(* IEC 61131-3 sources: SRCI_CLIENT_PLC/RobotLibrary/Library/POUs/Read/MC_ReadActualTCPVelocity/Structures, 4 files *)

(* ---- ReadActualTCPVelocityOutCmd.st ---- *)
{attribute 'pack_mode' := '1'}
// -------------------------------------------------------------------------
//  SRCI Robot Library
// -------------------------------------------------------------------------
//
//  Object:      ReadActualTCPVelocityOutCmd
//  Author:      Thorsten Brach
//  Date:        2024-08-09
//
//  Description:
//
//
//  Copyright:
//    (C) 2024 Thorsten Brach. All rights reserved
//             Licensed under the MIT License.
//
//  Disclaimer:
//    This project is provided without any guarantee and can be used for
//    private and commercial purposes. Any use is at the user’s
//    own risk and responsibility.
//
// -------------------------------------------------------------------------
TYPE ReadActualTCPVelocityOutCmd :
STRUCT
  /// Absolute actual velocity of the robot’s TCP. [mm/s]
  ActualTCPVelocity  : REAL;
  /// Index of tool of returned velocity
  /// •      0: Flange
  /// • 1..254: Tool frames
  ToolNoReturn       : USINT;
  /// Index of frame of returned position
  /// •      0: WCS
  /// • 1..254: User frames
  FrameNoReturn      : USINT;
  /// Unique system-generated ID of the "Action" when the function is triggered
  /// • >0: The "Action" is started by the trigger function with identical FollowID.
  /// • <0: The "Action" is stopped by the trigger function with identical FollowID.
  /// For more information see chapter 5.5.12.4
  OriginID           : INT;
  /// Relates to ListenerID >0 Number of successful trigger -based command invocations
  /// For more information refer to chapter 5.5.12.4
  InvocationCounter  : USINT;
END_STRUCT
END_TYPE

(* ---- ReadActualTCPVelocityParCmd.st ---- *)
{attribute 'pack_mode' := '1'}
// -------------------------------------------------------------------------
//  SRCI Robot Library
// -------------------------------------------------------------------------
//
//  Object:      ReadActualTCPVelocityParCmd
//  Author:      Thorsten Brach
//  Date:        2024-08-09
//
//  Description:
//
//
//  Copyright:
//    (C) 2024 Thorsten Brach. All rights reserved
//             Licensed under the MIT License.
//
//  Disclaimer:
//    This project is provided without any guarantee and can be used for
//    private and commercial purposes. Any use is at the user’s
//    own risk and responsibility.
//
// -------------------------------------------------------------------------
TYPE ReadActualTCPVelocityParCmd :
STRUCT
  /// Index of tool of returned velocity
  /// •      0: Flange (default)
  /// • 1..254: Tool frames
  ToolNo             : USINT;
  /// Index of frame
  /// •      0: WCS (default)
  /// • 1..254: User frames
  FrameNo            : USINT;
  /// ID of associated trigger function
  /// •  0: No Trigger (default) -> No trigger related behavior
  /// • >0: Trigger              -> Start executing when the trigger function with the identical EmitterID is triggered.
  /// Always positive. For more information, see chapter 5.5.12 Triggers
  ListenerID         : SINT;
END_STRUCT
END_TYPE

(* ---- ReadActualTCPVelocityRecvData.st ---- *)
{attribute 'pack_mode' := '1'}
// -------------------------------------------------------------------------
//  SRCI Robot Library
// -------------------------------------------------------------------------
//
//  Object:      ReadActualTCPVelocityRecvData
//  Author:      Thorsten Brach
//  Date:        2024-08-09
//
//  Description:
//
//
//  Copyright:
//    (C) 2024 Thorsten Brach. All rights reserved
//             Licensed under the MIT License.
//
//  Disclaimer:
//    This project is provided without any guarantee and can be used for
//    private and commercial purposes. Any use is at the user’s
//    own risk and responsibility.
//
// -------------------------------------------------------------------------
TYPE ReadActualTCPVelocityRecvData EXTENDS RspHeader :
STRUCT
  /// Relates to ListenerID >0
  /// Number of successful trigger-based command invocations - For more information refer TO chapter 5.5.12.4
  InvocationCounter : USINT;
  /// Reserve
  Reserve           : SINT;
  /// Unique system-generated ID of the "Action" when the function is triggered.
  /// • >0: The "Action" is started by the trigger funcrion with identical FollowID.
  /// • <0: The "Action" is stopped by the trigger function with identical FollowID.
  /// For more information see chapter 5.5.12.4 EmitterID, ListenerID, FollowID and OriginID
  OriginID          : INT;
  /// Absolute actual velocity of the robot’s TCP. [mm/s]
  ActualTCPVelocity  : REAL;
  /// Index of tool of returned velocity
  /// •      0: Flange
  /// • 1..254: Tool frames
  ToolNoReturn       : USINT;
  /// Index of frame of returned position
  /// •      0: WCS
  /// • 1..254: User frames
  FrameNoReturn      : USINT;
END_STRUCT
END_TYPE

(* ---- ReadActualTCPVelocitySendData.st ---- *)
{attribute 'pack_mode' := '1'}
// -------------------------------------------------------------------------
//  SRCI Robot Library
// -------------------------------------------------------------------------
//
//  Object:      ReadActualTCPVelocitySendData
//  Author:      Thorsten Brach
//  Date:        2024-08-09
//
//  Description:
//
//
//  Copyright:
//    (C) 2024 Thorsten Brach. All rights reserved
//             Licensed under the MIT License.
//
//  Disclaimer:
//    This project is provided without any guarantee and can be used for
//    private and commercial purposes. Any use is at the user’s
//    own risk and responsibility.
//
// -------------------------------------------------------------------------
TYPE ReadActualTCPVelocitySendData EXTENDS CmdHeader:
STRUCT
  /// Index of tool of returned velocity
  /// •      0: Flange (default)
  /// • 1..254: Tool frames
  ToolNo             : USINT;
  /// Index of frame
  /// •      0: WCS (default)
  /// • 1..254: User frames
  FrameNo            : USINT;
END_STRUCT
END_TYPE
